// TIA Portal V19 export
DATA_BLOCK "Tacho2_EM03"   // DB4
VERSION : 1.0
// stored: InstanceOfName EM03_Alimentacion, InstanceOfType FB
"EM03_Alimentacion"
   // VAR_INPUT
   //    In : "EM03_Input";
   //    FeedPV : Real;
   // END_VAR
   // VAR_OUTPUT
   //    Out : "EM03_Output";
   //    CM_PIC_MV : Real;
   //    CM_Vlv_MP_Out : Array[1..2] of Bool;
   //    CM_Agua_Out : Real;
   //    SensorAlarm : Bool;
   //    CMAlarm : Bool;
   // END_VAR
   // VAR
   //    State : Int;
   //    ActiveAction : Int;
   //    AlarmLatched : Bool;
   //    FaultCode : Int;
   //    TimerStable { S7_SetPoint := 'True'} : TON_TIME;
   //    TrigStart { S7_SetPoint := 'True'} : R_TRIG;
   //    TrigStop { S7_SetPoint := 'True'} : R_TRIG;
   //    TrigHold { S7_SetPoint := 'True'} : R_TRIG;
   //    TrigAbort { S7_SetPoint := 'True'} : R_TRIG;
   //    TrigReset { S7_SetPoint := 'True'} : R_TRIG;
   //    CM_PIC_Feed { S7_SetPoint := 'True'} : "PidL";
   //    CM_Vlv_MateriaPrima { S7_SetPoint := 'True'} : Array[1..2] of "VlvL";
   //    CM_Vlv_Agua { S7_SetPoint := 'True'} : "OpAn";
   // END_VAR
BEGIN
   In.FeedSP := 50.0;
   In.WashSP := 20.0;
   CM_PIC_Feed.DataHMI.identName := 'LCV-212';
   CM_PIC_Feed.DataHMI.comment := 'Nivel';
   CM_Vlv_MateriaPrima[1].DataHMI.identName := 'XSV112A';
   CM_Vlv_MateriaPrima[2].DataHMI.identName := 'XSV112B';
   CM_Vlv_MateriaPrima[1].DataHMI.comment := 'Melad.Clara';
   CM_Vlv_MateriaPrima[2].DataHMI.comment := 'Melad.Cruda';
END_DATA_BLOCK
